# EPICS substitutions: db/Beckhoff_6XXX/ecmcEL6688.substitutions
file "ecmcEL6688.template"
{
  pattern {}
          {}
}
